Staubli VAL3: showActive.pgx

program showActive(num x_nIndex)
begin
  bActive=(safeTemp:sSPoint[x_nIndex].bActive==true)
end
